FUNCTION_BLOCK FB_MeanValue
VAR_INPUT
	(* Input variables / Eingang Variablen *)
	bEnable					:BOOL;						(* Enable FB signal *)
	bReset					:BOOL;						(* Reset measurement *)
	bExecute				:BOOL;						(* Execute measurement *)
	bAbort					:BOOL;						(* Abort measurement *)
	lrSampleValue			:LREAL;						(* Sample measurement value *)
	lrSampleValueMin		:LREAL;						(* Sample measurement value minimum *)
	lrSampleValueMax		:LREAL;						(* Sample measurement value maximum *)
	udnSampleTime			:UDINT := 100;				(* Sample time [ms] *)
	udnSampleDeathStart		:UDINT;						(* Amount of death sample from start *)
	tMaxTime				:TIME := T#1092M;			(* Maximum time *)
END_VAR
VAR_OUTPUT
	(* Output variables / Ausgang Variablen *)
	lrMeanValue				:LREAL;						(* Mean measurement value *)
END_VAR
VAR_IN_OUT

END_VAR
VAR
	(* Enummerations *)

	(* Variables *)
	udnCounter				:UDINT;
	lrTotalValue			:LREAL;						(* Total measurement value *)
	bFirstTime				:BOOL;

	(* References *)

	(* Interfaces *)

	(* Instances *)
	fbCycleTime					:FB_Timer;
	
END_VAR

IF NOT bEnable
THEN
	lrMeanValue := lrSampleValue;
	bFirstTime := FALSE;
	RETURN;
END_IF;

IF NOT bFirstTime
THEN

	bFirstTime := TRUE;
END_IF;

(* Measuring time of cycle *)
fbCycleTime(
	bEnable := TRUE,
	bReset := bReset,
	bStartStop := bExecute,
	bStop := NOT bExecute OR bAbort,
	tMaxTime := tMaxTime
);

IF fbCycleTime.bTimeStarted 
THEN
	IF fbCycleTime.stActTime.dwMiliSec >= udnSampleTime * udnCounter
	THEN
		IF (lrSampleValue > lrSampleValueMin
			AND lrSampleValue < lrSampleValueMax)
			OR lrSampleValueMin = lrSampleValueMax
		THEN
			udnCounter := udnCounter + 1;
			
			IF udnCounter > udnSampleDeathStart
			THEN
				lrTotalValue := lrTotalValue + lrSampleValue;		
				lrMeanValue := lrTotalValue / UDINT_TO_LREAL(udnCounter - udnSampleDeathStart);
			END_IF
		END_IF		
	END_IF
ELSE
	lrTotalValue := 0;
	udnCounter := 0;
END_IF

END_FUNCTION_BLOCK

(* stored: Version 1.1.0.1, ProductVersion 3.1.4024.15
   POU FB_MeanValue: Id {8e30639c-70f9-46ab-b3d1-d9017ceae5a2}, SpecialFunc None *)
